// CONVERTE TIME IN SECONDI (REAL)
FUNCTION F_TimeToSeconds : REAL
VAR_INPUT
	tTime	:	TIME;
END_VAR
VAR
END_VAR

F_TimeToSeconds	:=	TIME_TO_REAL(tTime) * GVL_Conversions.TIME_TO_SECONDS;

END_FUNCTION

(* stored: Version 1.1.0.1, ProductVersion 3.1.4024.9
   POU F_TimeToSeconds: Id {8320d3a7-89fe-4fcd-accd-72e89d860407}, SpecialFunc None *)
